// TIA Portal V19 export
// export: Created 2026-11-08T08:30:00.0000000Z, ExportSetting WithReadOnly
TYPE "UDT_ExampleCfg"
   STRUCT
      Enable : Bool;
      Delay : Time := T#5S;
   END_STRUCT;
END_TYPE
